// TIA Portal V21 export
// export: Created 2026-11-10T07:35:01.528894Z, ExportSetting WithDefaults, DisplayName Totally Integrated Automation Portal, DisplayVersion V21 Update 3, DisplayName STEP 7 Professional, DisplayVersion V21 Update 3, DisplayName STEP 7 Safety, DisplayVersion V21, DisplayName Tech WebApplication, DisplayVersion V21, DisplayName WinCC Basic/Comfort/Advanced, DisplayVersion V21 Update 3, DisplayName WinCC Unified, DisplayVersion V21 Update 3
FUNCTION_BLOCK "FB_Lad_ex009"   // FB8, LAD
{ S7_Optimized_Access := 'TRUE' }
VERSION : 0.1
// stored: AutoNumber true, IsIECCheckEnabled false, IsRetainMemResEnabled false, MemoryReserve 100, SetENOAutomatically false, UDAEnableTagReadback false
   VAR_INPUT
      v_ret_val : Int;
   END_VAR
   VAR_OUTPUT
      v_out : DTL;
   END_VAR
BEGIN

REGION Network 1: RD_LOC_T - Read local time
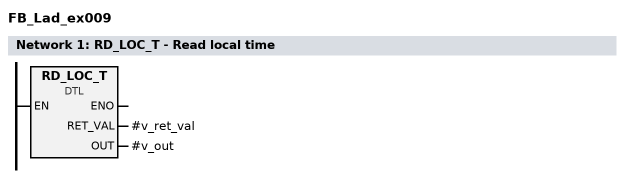
   RUNG wire#powerrail
      { S7_Templates := "date_type := DTL" } RD_LOC_T(RET_VAL => #v_ret_val, OUT => #v_out)
   END_RUNG
   // the same network as SCL:
   #v_ret_val := RD_LOC_T(OUT => #v_out);
END_REGION
END_FUNCTION_BLOCK
